(* IEC 61131-3 sources: PortalRobot/Portal_robot/Device/application/ST/ST_AXIS, 10 files *)

(* ---- E_AXIS_STATE.st ---- *)
{attribute 'qualified_only'}
{attribute 'strict'}
TYPE E_AXIS_STATE :
(
	DISABLED,
	POWERING,
	POWERING_DOWN,
	READY,
	JOGGING,
	JOG_DECELERATING,
	HOMING,
	MOVE_ABSOLUTE,
	MOVE_RELATIVE,
	STOPPING,
	STOP_RELEASE,
	ERROR_RESET_MANAGER,
	RESET_AXIS_ERROR,
	RESET_RELEASE,
	RESET_FINISH
);
END_TYPE

(* ---- ST_AXIS.st ---- *)
TYPE ST_AXIS :
STRUCT
	Command     : ST_AXIS_COMMANDS; // Команды оси
	Status      : ST_AXIS_STATUS; // Рабочие статусы оси
	Diag        : ST_AXIS_DIAGNOSTICS; // Состояние автомата и текстовая диагностика
	Error       : ST_AXIS_ERROR_CODES; // Активные и последние ошибки
	MotionParam : ST_AXIS_MOTION_PARAMS; // Параметры движения
	Timeouts    : ST_AXIS_TIMEOUTS; // Допустимое время выполнения шагов

END_STRUCT
END_TYPE

(* ---- ST_AXIS_COMMANDS.st ---- *)
TYPE ST_AXIS_COMMANDS :
STRUCT
    xEnable            : BOOL; // Импульс запроса включения оси
    xDisable           : BOOL; // Импульс запроса отключения оси
	xGlobalError       : BOOL; // Глобальная ошибка ячейки
	xPowerPermit       : BOOL; // Разрешение подачи питания на привод
    xResetAllError     : BOOL; // Общий сброс ошибок оси
    xResetAxisError    : BOOL; // Сброс ошибок привода и SoftMotion
    xResetLogicalError : BOOL; // Сброс логических ошибок блока
    xStop              : BOOL; // Команда контролируемой остановки
    xHome              : BOOL; // Команда поиска домашней позиции
    xMoveAbsolute      : BOOL; // Команда абсолютного перемещения
    xMoveRelative      : BOOL; // Команда относительного перемещения
    xJogPositive       : BOOL; // Толчковое движение в положительном направлении
    xJogNegative       : BOOL; // Толчковое движение в отрицательном направлении
END_STRUCT
END_TYPE

(* ---- ST_AXIS_DIAGNOSTICS.st ---- *)
TYPE ST_AXIS_DIAGNOSTICS :
STRUCT
    iStep            : E_AXIS_STATE; // Текущий шаг автомата оси
    iLastErrorStep   : INT; // Шаг, на котором возникла последняя ошибка
    sStepName        : STRING[80]; // Текстовое имя текущего шага
    sWaitReason      : STRING[120]; // Причина ожидания на текущем шаге
    sErrorText       : STRING[120]; // Текст активной ошибки
    sWarningText     : STRING[120]; // Текст активного предупреждения
    stWarning        : ST_WARNING_EVENT; // Последнее предупреждение оси для общего журнала
    tStepElapsed     : TIME; // Время нахождения на текущем шаге
    tStepPreset      : TIME; // Допустимое время текущего шага
    xStepTimeout     : BOOL; // Превышено допустимое время шага
    udiActualErrorID : UDINT; // Код активной ошибки
    udiLastErrorID   : UDINT; // Код последней ошибки
END_STRUCT
END_TYPE

(* ---- ST_AXIS_ERROR.st ---- *)
TYPE ST_AXIS_ERROR :
STRUCT
	MC_POWER_ERROR       : BOOL; // Ошибка MC_Power
	MC_RESET_ERROR       : BOOL; // Ошибка MC_Reset
	MC_STOP_ERROR        : BOOL; // Ошибка MC_Stop
	MC_JOG_ERROR         : BOOL; // Ошибка MC_Jog
	MC_HOME_ERROR        : BOOL; // Ошибка MC_Home
	MC_MOVE_ABS_ERROR    : BOOL; // Ошибка MC_MoveAbsolute
	MC_MOVE_REL_ERROR    : BOOL; // Ошибка MC_MoveRelative
	READ_POSITION_ERROR  : BOOL; // Ошибка чтения позиции
	READ_STATUS_ERROR    : BOOL; // Ошибка чтения статуса оси
	AXIS_ERRORSTOP       : BOOL; // Ось находится в ErrorStop
	FB_ERROR_OCCURRED    : BOOL; // SoftMotion сообщил внутреннюю ошибку
	COMMAND_ABORTED      : BOOL; // Команда движения была прервана
	UNKNOWN_AXIS_ERROR   : BOOL; // Неизвестная ошибка оси
	DRIVE_AXIS_ERROR     : BOOL; // Ошибка привода оси
	POWER_FEEDBACK_LOST  : BOOL; // Потеря силовой готовности при активной команде питания
	POWER_PERMIT_LOST    : BOOL; // Потеря разрешения питания
	GLOBAL_DURING_POWER  : BOOL; // Глобальная ошибка при включении
	GLOBAL_DURING_READY  : BOOL; // Глобальная ошибка в готовности
	GLOBAL_DURING_MOTION : BOOL; // Глобальная ошибка во время движения
	JOG_CONFLICT         : BOOL; // Одновременно поданы Jog+ и Jog-
	MOVE_ABS_NOT_HOMED   : BOOL; // Абсолютное движение без Home
	MOVE_REL_NOT_HOMED   : BOOL; // Относительное движение без Home
	STEP_TIMEOUT         : BOOL; // Превышено время выполнения шага
	UNKNOWN_STEP         : BOOL; // Неизвестное состояние автомата
END_STRUCT
END_TYPE

(* ---- ST_AXIS_ERROR_CODES.st ---- *)
TYPE ST_AXIS_ERROR_CODES :
STRUCT
    dwAxisErrorActual     : DWORD; // Текущие ошибки блоков SoftMotion
    dwAxisErrorLatched    : DWORD; // Защёлкнутые ошибки SoftMotion
    dwAxisError           : DWORD; // Общая активная маска ошибок оси
    dwAxisErrorLast       : DWORD; // Последняя ненулевая маска ошибок оси
    dwDriveAxisErrorID    : DWORD; // Код ошибки привода
    dwLogicalErrorLatched : DWORD; // Защёлкнутые логические ошибки
    dwLogicalError        : DWORD; // Общая активная маска логических ошибок
    dwLogicalErrorLast    : DWORD; // Последняя ненулевая маска логических ошибок
    dwWarningLatched      : DWORD; // Защёлкнутые предупреждения
    dwWarning             : DWORD; // Активные предупреждения
    dwAllError            : DWORD; // Сводная маска ошибок
    dwAlarmActive         : DWORD; // Собственные аварии оси для общего журнала
    stErrorActive         : ST_AXIS_ERROR; // Расшифровка активных ошибок
    stErrorLast           : ST_AXIS_ERROR; // Расшифровка последних ошибок
END_STRUCT
END_TYPE

(* ---- ST_AXIS_FAULT_REQUEST.st ---- *)
TYPE ST_AXIS_FAULT_REQUEST :
STRUCT
	xEnabled     : BOOL; // Глобальное разрешение диагностической инъекции
	xJogConflict : BOOL; // Импульс одновременного запроса Jog+ и Jog-
END_STRUCT
END_TYPE

(* ---- ST_AXIS_MOTION_PARAMS.st ---- *)
TYPE ST_AXIS_MOTION_PARAMS :
STRUCT
    lrTargetPosition : LREAL; // Целевая абсолютная позиция
    lrDistance       : LREAL; // Дистанция относительного перемещения
    lrHomePosition   : LREAL; // Координата домашней позиции
    lrVelocity       : LREAL; // Скорость движения
    lrAcceleration   : LREAL; // Ускорение
    lrDeceleration   : LREAL; // Замедление
    lrJerk           : LREAL; // Рывок
END_STRUCT
END_TYPE

(* ---- ST_AXIS_STATUS.st ---- *)
TYPE ST_AXIS_STATUS :
STRUCT
	xStandstill : BOOL; // MC_ReadStatus: подтверждённый останов, включая Disabled/ErrorStop
    xPowered            : BOOL; // На привод подано питание
	xPowerStageOn        : BOOL; // Фактическое подтверждение включения силовой части
	xDriveStartOn        : BOOL; // Фактическое подтверждение снятого QuickStop
	xPowerOff            : BOOL; // Силовая часть отключена и QuickStop активен
    xBusy               : BOOL; // Ось выполняет команду
    xDone               : BOOL; // Последняя команда завершена
    xError              : BOOL; // Активна любая ошибка оси
    xHomed              : BOOL; // Ось прошла поиск домашней позиции
    xLocalError         : BOOL; // Активна внутренняя ошибка блока
    xMotionBusy         : BOOL; // Активен один из блоков движения
    xCanStartMotion     : BOOL; // Разрешён запуск новой команды движения
    xAxisError          : BOOL; // Активна ошибка привода или SoftMotion
    xLogicalError       : BOOL; // Активна логическая ошибка блока
    xWarning            : BOOL; // Активно предупреждение
    xAxisResetNeeded    : BOOL; // Требуется сброс ошибки привода
    xLogicalResetNeeded : BOOL; // Требуется сброс логической ошибки
	lrActualPosition    : REAL; // Текущая позиция оси
END_STRUCT
END_TYPE

(* ---- ST_AXIS_TIMEOUTS.st ---- *)
TYPE ST_AXIS_TIMEOUTS :
STRUCT
	xDisableOnError : BOOL := TRUE; // Отключать привод при логической ошибке
    tPowerFeedbackLossTimeout : TIME := T#500MS; // Потеря силовой готовности при сохраняющемся запросе питания
    tPowerTimeout   : TIME := T#5S; // Время ожидания включения или отключения питания
    tResetTimeout   : TIME := T#5S; // Время ожидания сброса ошибки
    tStopTimeout    : TIME := T#5S; // Время ожидания остановки
    tHomeTimeout    : TIME := T#30S; // Время ожидания поиска домашней позиции
    tMoveTimeout    : TIME := T#15S; // Время ожидания завершения перемещения
END_STRUCT
END_TYPE
